Fanuc KAREL source: KA00092.KL

PROGRAM KA00092
%NOLOCKGROUP
VAR
  SRC: JOINTPOS
  DST: JOINTPOS
BEGIN
  DST = SRC
END KA00092
